RoboDK station: drawbot.rdk

Station DrawBot (saved by RoboDK 6.0.7). Poses are relative to the parent item; angles as X-Y-Z fixed-axis rotations.
Station parameters (name, value as stored): WB_WIDTH_MM, 335.73, WB_HEIGHT_MM, 293.87, DRAWBOT_HOME_SEED, [221.439, -65.915, 102.122, -158.595, -78.539, -31.343]
